(* IEC 61131-3 sources: plcassist-cli/packages/volt-lsp-iec/test-corpus/awa-palletizer/Device/Plc Logic/Application/Library Manager/VisuShared, 17 files *)

(* ---- EVENT_SYNC_FILE.gvl ---- *)
VAR_GLOBAL
	EVT_SYNCFILETRANSFER : UDINT := 16#10002;
	CMPID_CMPFILETRANSFER : UDINT := 16#5E;
	SYNCFILE_TYPE_START : UINT := 1;
	SYNCFILE_TYPE_END : UINT := 2;
END_VAR

(* ---- VISUSHARED_GLOBALS.gvl ---- *)
VAR_GLOBAL
	G_SYNCFILETRANSFEREVENT : Visu_FbSyncFileTransferEvent;
	G_UILOADTEXTLIST : UDINT;
	G_UILOADTEXTLISTOCBIT : UDINT := 0;
	G_UILOADTEXTLISTBEFOREOCBIT : UDINT := 1;
	G_UILOADTEXTLISTDLBIT : UDINT := 2;
	G_DATETIMEPROVIDER : Visu_FbDateTimeProvider;
END_VAR

(* ---- ICALLONINITIALIZEBASE.itf ---- *)
INTERFACE ICALLONINITIALIZEBASE
END_INTERFACE

METHOD INIT : BOOL
END_METHOD

(* ---- CONVERTDATETIME.fun ---- *)
FUNCTION CONVERTDATETIME : ULINT
VAR_INPUT
	UIYEAR : YEAR;
END_VAR
VAR_OUTPUT
	EERRORID : ERROR;
END_VAR
VAR_IN_OUT
	DTDATETIME : DateTime;
END_VAR
END_FUNCTION

(* ---- EXTRACTYEARMONTHDAY.fun ---- *)
FUNCTION EXTRACTYEARMONTHDAY : ERROR
VAR_INPUT
	ULIDATETIME : ULINT;
END_VAR
VAR_OUTPUT
	UIYEAR : YEAR;
	UIMONTH : MONTH;
	UIDAY : DAY;
END_VAR
END_FUNCTION

(* ---- GETLIBVERSION.fun ---- *)
FUNCTION GETLIBVERSION : VERSION
END_FUNCTION

(* ---- GETLIBVERSIONNUMBER.fun ---- *)
FUNCTION GETLIBVERSIONNUMBER : DWORD
END_FUNCTION

(* ---- GETTASKBYNAME.fun ---- *)
FUNCTION GETTASKBYNAME : BOOL
VAR_INPUT
	SZAPPNAME : STRING(CmpApp.GlobalConstants.MAX_LEN_APPLNAME);
	SZTASK : POINTER TO STRING;
END_VAR
VAR_OUTPUT
	HTASK : RTS_IEC_HANDLE;
END_VAR
END_FUNCTION

(* ---- ISLIBRELEASED.fun ---- *)
FUNCTION ISLIBRELEASED : BOOL
END_FUNCTION

(* ---- ISTASKRUNNING.fun ---- *)
FUNCTION ISTASKRUNNING : BOOL
VAR_INPUT
	HTASK : RTS_IEC_HANDLE;
	SZAPPNAME : STRING(CmpApp.GlobalConstants.MAX_LEN_APPLNAME);
END_VAR
END_FUNCTION

(* ---- LEAPYEARS.fun ---- *)
FUNCTION LEAPYEARS : UINT
VAR_INPUT
	UISTARTYEAR : YEAR;
	UIENDYEAR : YEAR;
END_VAR
VAR_OUTPUT
	EERRORID : ERROR;
END_VAR
END_FUNCTION

(* ---- LOADTEXTLISTBEFOREONLINECHANGE.fun ---- *)
FUNCTION LOADTEXTLISTBEFOREONLINECHANGE : BOOL
END_FUNCTION

(* ---- RELOADTEXTLISTSIFNECESSARY.fun ---- *)
FUNCTION RELOADTEXTLISTSIFNECESSARY : BOOL
VAR_INPUT
	BDOWNLOAD : BOOL;
	BFORCE : BOOL;
END_VAR
END_FUNCTION

(* ---- UTILTIMEZONELOCALTOUTC.fun ---- *)
FUNCTION UTILTIMEZONELOCALTOUTC : SYSTIME
VAR_INPUT
	ULILOCALTIME : SYSTIME;
END_VAR
VAR_OUTPUT
	EERRORID : ERROR;
	EPERIOD : PERIOD;
END_VAR
VAR_IN_OUT
	TZTIMEZONE : TimeZone;
END_VAR
END_FUNCTION

(* ---- VISU_FBDATETIMEPROVIDER.fb ---- *)
FUNCTION_BLOCK VISU_FBDATETIMEPROVIDER
VAR_INPUT
	ENDATETIMELIBRARY : VisuEnumDateTimeLibrary := VisuEnumDateTimeLibrary.UseSysTimeRTC;
	TZTIMEZONE : Util.TimeZone;
END_VAR
END_FUNCTION_BLOCK

METHOD CONVERTLOCALTOUTCTIME : SYSTIME
VAR_INPUT
	LOCALTIME : SYSTIME;
END_VAR
VAR_OUTPUT
	EERRORID : ERROR;
	IUTCOFFSET : INT;
END_VAR
END_METHOD

METHOD CONVERTUTCTOLOCALTIME : SYSTIME
VAR_INPUT
	UTCTIME : SYSTIME;
END_VAR
VAR_OUTPUT
	EERRORID : ERROR;
	IUTCOFFSET : INT;
END_VAR
END_METHOD

METHOD GETCURRENTLOCALTIME : SYSTIME
VAR_OUTPUT
	EERRORID : ERROR;
	IUTCOFFSET : INT;
END_VAR
END_METHOD

METHOD GETCURRENTUTCTIME : SYSTIME
VAR_OUTPUT
	EERRORID : ERROR;
END_VAR
END_METHOD

(* ---- VISU_FBINITONSTARTUP.fb ---- *)
FUNCTION_BLOCK VISU_FBINITONSTARTUP
VAR
	_ARR : ARRAY [0..(MAX_STARTUPINITIALZATIONS - 1)] OF ICallOnInitializeBase;
	_ICOUNT : INT;
	MAX_STARTUPINITIALZATIONS : INT := 5;
END_VAR
END_FUNCTION_BLOCK

METHOD CALLINITIALIZE
END_METHOD

METHOD REGISTER : BOOL
VAR_INPUT
	INSTANCE : ICallOnInitializeBase;
END_VAR
END_METHOD

(* ---- VISU_FBSYNCFILETRANSFEREVENT.fb ---- *)
FUNCTION_BLOCK VISU_FBSYNCFILETRANSFEREVENT
VAR
	_HEVENTSTART : SysTypes.RTS_IEC_HANDLE := SysTypes.RTS_INVALID_HANDLE;
	_HINTERFACESTART : SysTypes.RTS_IEC_HANDLE := SysTypes.RTS_INVALID_HANDLE;
	_ITFEVENTCALLBACK : CmpEventMgr_Interfaces.ICmpEventCallback;
END_VAR
END_FUNCTION_BLOCK

METHOD EVENTCALLBACK : SysTypes.RTS_IEC_RESULT
VAR_INPUT
	PEVENTPARAM : POINTER TO EventParam;
END_VAR
END_METHOD

METHOD FB_EXIT : BOOL
VAR_INPUT
	BINCOPYCODE : BOOL;
END_VAR
END_METHOD

METHOD FB_INIT : BOOL
VAR_INPUT
	BINITRETAINS : BOOL;
	BINCOPYCODE : BOOL;
END_VAR
END_METHOD
